// TIA Portal V19 export
// export: Created 2026-10-19T00:00:00.0000000Z, ExportSetting None
FUNCTION_BLOCK "FB_ProbeFbd"   // FB1, FBD
TITLE = FB_ProbeFbd
{ S7_Optimized_Access := 'TRUE' }
// FBD FB_ProbeFbd → FBD (c2s7)
// stored: AutoNumber true, MemoryReserve 100, SetENOAutomatically false
   VAR_INPUT
      rLevel : Real;
      rHigh : Real;
      xEnable : Bool;
      xAck : Bool;
   END_VAR
   VAR_OUTPUT
      xOut : Bool;
   END_VAR
   VAR
      xHigh : Bool;
      xAlarm : Bool;
   END_VAR
BEGIN

REGION Network 1
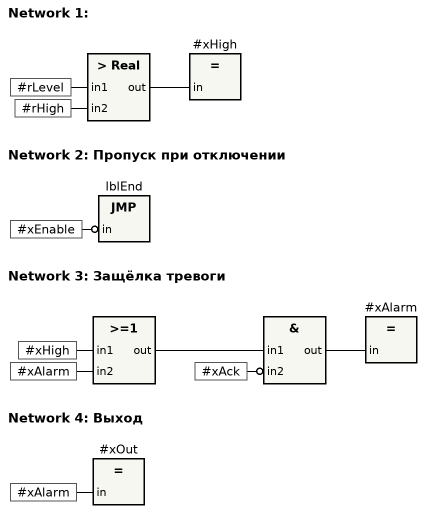
   #xHigh := #rLevel > #rHigh;
END_REGION

REGION Network 2: Пропуск при отключении
   IF NOT #xEnable THEN GOTO <??.?>; END_IF;
END_REGION

REGION Network 3: Защёлка тревоги
   #xAlarm := (#xHigh OR #xAlarm) AND NOT #xAck;
END_REGION

REGION Network 4: Выход
   lblEnd:
   #xOut := #xAlarm;
END_REGION
END_FUNCTION_BLOCK
